(* Schneider Machine Expert - Basic project subroutine_sr0_watch3, file version 3.0.0.0 *)
(* ProjectInformations: Name=New project *)

HARDWARE
  Cpu 0: TM200CE40T
  EthernetConfiguration: NetworkName=M200, IpAllocationMode=FixedAddress, IpAddress=0.0.0.0, SubnetMask=0.0.0.0
  SerialLineConfiguration: Baud=Baud19200, Parity=ParityEven, DataBits=DataBits8, StopBits=StopBits1, PhysicalMedium=PhysicalMediumRs485, TransmissionMode=TransmissionModeModbusRtu, SlaveId=1, Addressing=SlaveAddressing
  MastTask: UsePeriodScanMode=false, PeriodScan=100
  FastTask: Period=255
  CpuBehavior: StartingMode=StartAsPreviousState, AutoSaveRamOnEeprom=true, WatchdogPeriod=250

SYMBOLS  (address, symbol, comment, settings)

POU New POU
  (* SectionNumber=0 *)

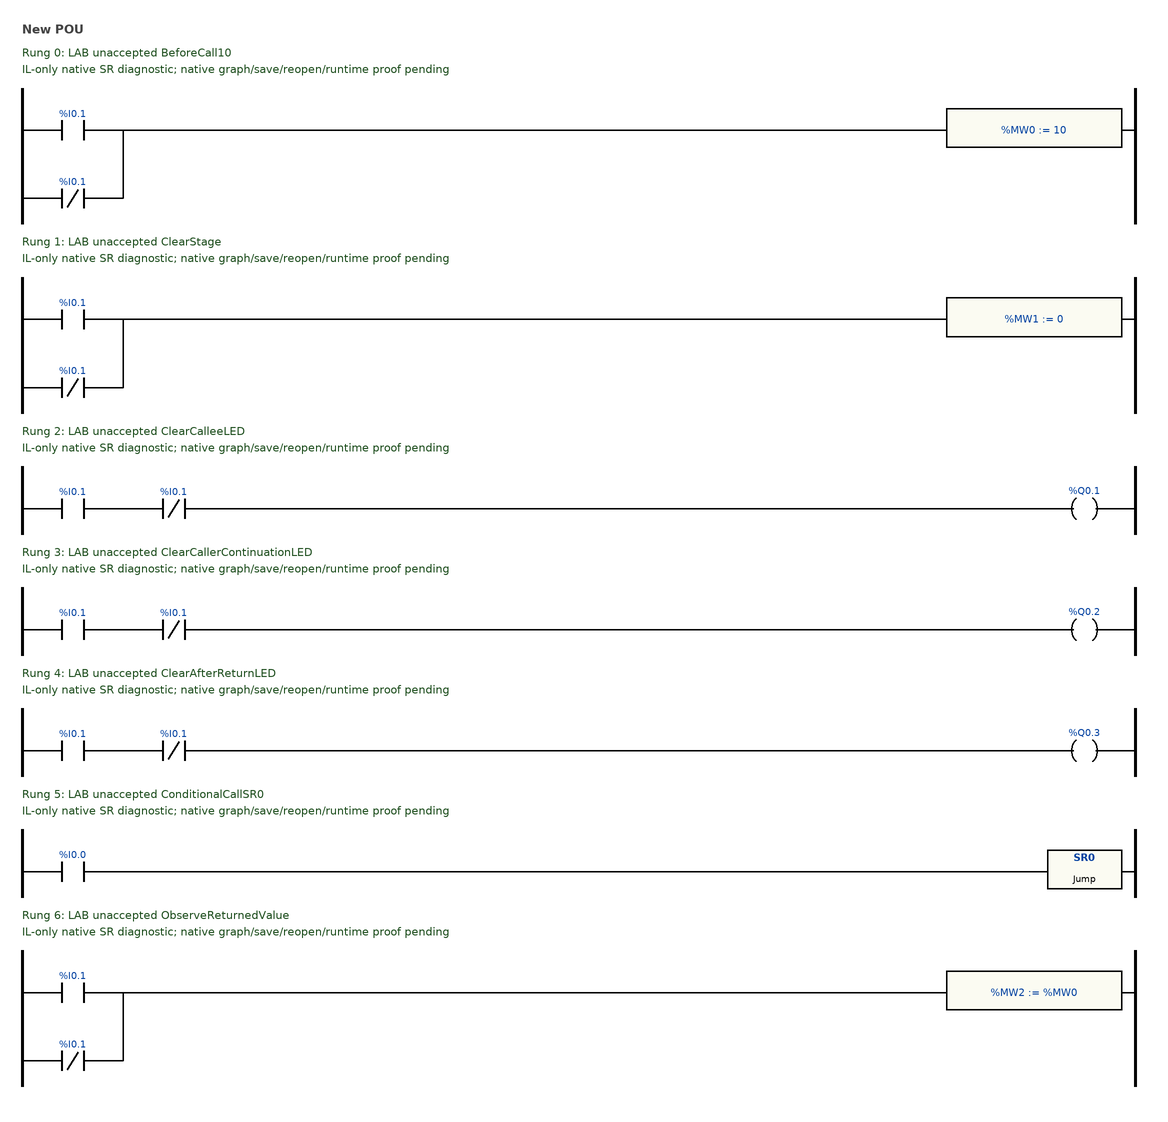

// Rung 0: LAB unaccepted BeforeCall10
// IL-only native SR diagnostic; native graph/save/reopen/runtime proof pending
  LD %I0.1
  ORN %I0.1
  [ %MW0 := 10 ]
  // as ST:
  //   IF %I0.1 OR NOT %I0.1 THEN %MW0 := 10; END_IF;

// Rung 1: LAB unaccepted ClearStage
// IL-only native SR diagnostic; native graph/save/reopen/runtime proof pending
  LD %I0.1
  ORN %I0.1
  [ %MW1 := 0 ]
  // as ST:
  //   IF %I0.1 OR NOT %I0.1 THEN %MW1 := 0; END_IF;

// Rung 2: LAB unaccepted ClearCalleeLED
// IL-only native SR diagnostic; native graph/save/reopen/runtime proof pending
  LD %I0.1
  ANDN %I0.1
  ST %Q0.1
  // as ST:
  //   %Q0.1 := %I0.1 AND NOT %I0.1;

// Rung 3: LAB unaccepted ClearCallerContinuationLED
// IL-only native SR diagnostic; native graph/save/reopen/runtime proof pending
  LD %I0.1
  ANDN %I0.1
  ST %Q0.2
  // as ST:
  //   %Q0.2 := %I0.1 AND NOT %I0.1;

// Rung 4: LAB unaccepted ClearAfterReturnLED
// IL-only native SR diagnostic; native graph/save/reopen/runtime proof pending
  LD %I0.1
  ANDN %I0.1
  ST %Q0.3
  // as ST:
  //   %Q0.3 := %I0.1 AND NOT %I0.1;

// Rung 5: LAB unaccepted ConditionalCallSR0
// IL-only native SR diagnostic; native graph/save/reopen/runtime proof pending
  LD %I0.0
  SR0
  // as ST:
  //   IF %I0.0 THEN SR0(); END_IF;

// Rung 6: LAB unaccepted ObserveReturnedValue
// IL-only native SR diagnostic; native graph/save/reopen/runtime proof pending
  LD %I0.1
  ORN %I0.1
  [ %MW2 := %MW0 ]
  // as ST:
  //   IF %I0.1 OR NOT %I0.1 THEN %MW2 := %MW0; END_IF;

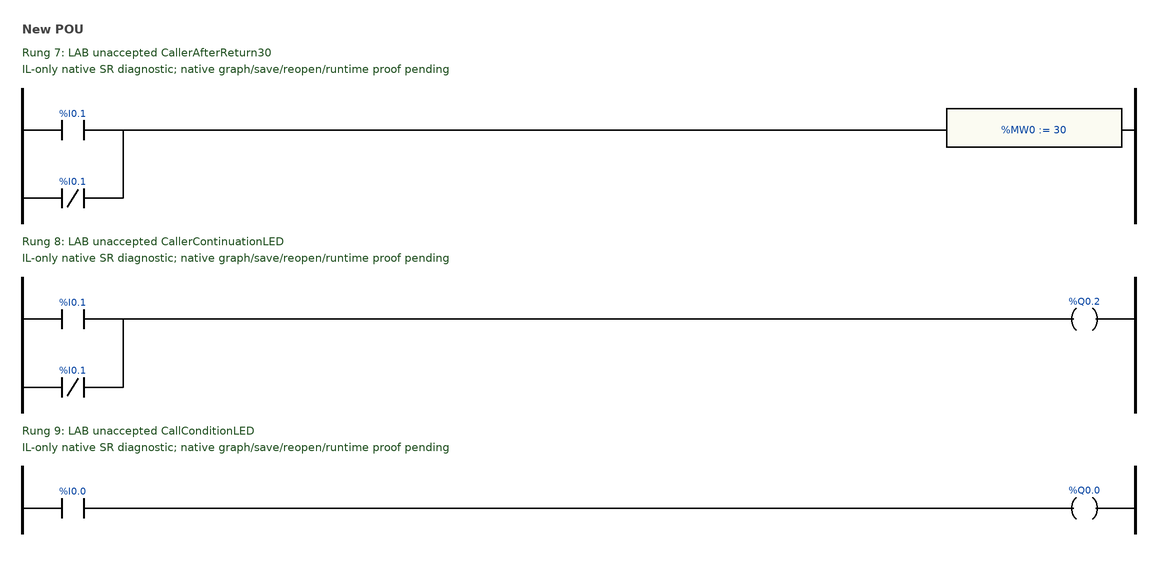

// Rung 7: LAB unaccepted CallerAfterReturn30
// IL-only native SR diagnostic; native graph/save/reopen/runtime proof pending
  LD %I0.1
  ORN %I0.1
  [ %MW0 := 30 ]
  // as ST:
  //   IF %I0.1 OR NOT %I0.1 THEN %MW0 := 30; END_IF;

// Rung 8: LAB unaccepted CallerContinuationLED
// IL-only native SR diagnostic; native graph/save/reopen/runtime proof pending
  LD %I0.1
  ORN %I0.1
  ST %Q0.2
  // as ST:
  //   %Q0.2 := %I0.1 OR NOT %I0.1;

// Rung 9: LAB unaccepted CallConditionLED
// IL-only native SR diagnostic; native graph/save/reopen/runtime proof pending
  LD %I0.0
  ST %Q0.0
  // as ST:
  //   %Q0.0 := %I0.0;

Subroutine LAB_SR0_LEAF
  (* SectionNumber=2, Number=0 *)

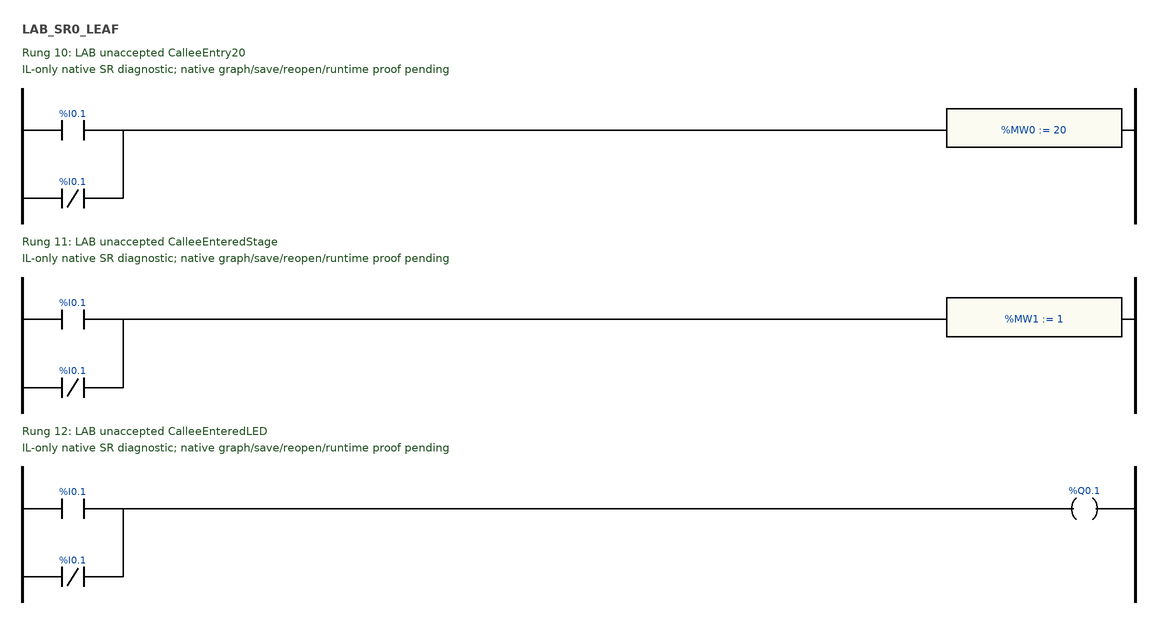

// Rung 10: LAB unaccepted CalleeEntry20
// IL-only native SR diagnostic; native graph/save/reopen/runtime proof pending
  LD %I0.1
  ORN %I0.1
  [ %MW0 := 20 ]
  // as ST:
  //   IF %I0.1 OR NOT %I0.1 THEN %MW0 := 20; END_IF;

// Rung 11: LAB unaccepted CalleeEnteredStage
// IL-only native SR diagnostic; native graph/save/reopen/runtime proof pending
  LD %I0.1
  ORN %I0.1
  [ %MW1 := 1 ]
  // as ST:
  //   IF %I0.1 OR NOT %I0.1 THEN %MW1 := 1; END_IF;

// Rung 12: LAB unaccepted CalleeEnteredLED
// IL-only native SR diagnostic; native graph/save/reopen/runtime proof pending
  LD %I0.1
  ORN %I0.1
  ST %Q0.1
  // as ST:
  //   %Q0.1 := %I0.1 OR NOT %I0.1;
